(* IEC 61131-3 sources: avi-aoi-management/scripts/ai-eval/ngau-nhien/kho/st-tt6-chon-bom-chinh/khung/src, 1 file *)

(* ---- ChonBomChinh.st ---- *)
FUNCTION_BLOCK ChonBomChinh
VAR_INPUT
    GIO_CHAY : ARRAY[1..4] OF UDINT;
    SAN_SANG : ARRAY[1..4] OF BOOL;
END_VAR
VAR_OUTPUT
    BOM : INT;
    THU_TU : ARRAY[1..4] OF INT;
END_VAR
    (* TODO: cài đặt theo đề bài *)
    BOM := 0;
END_FUNCTION_BLOCK
